(* IEC 61131-3 sources: plc-workbench/outputs/tia_32x4_20261108_results/tasks/15_PUBLIC_03/self_A/details/submissions/1/evaluation/formal, 1 file *)

(* ---- normalized.st ---- *)
FUNCTION_BLOCK Q03

   VAR_INPUT
      Value : REAL;
      hiLevel : REAL;
      loLevel : REAL;
      hystWindow : REAL;
   END_VAR
   VAR_OUTPUT
      hiAlarm : BOOL;
      loAlarm : BOOL;
      error : BOOL;
      status : WORD;
   END_VAR
   VAR
      valid : BOOL;
   END_VAR
VAR_INPUT
WBTEMP_0 : BOOL;
END_VAR

valid := WBTEMP_0;
   // Validity of configuration
   valid := FALSE;

   IF loLevel >= hiLevel THEN
      // Invalid limits: loLevel must be smaller than hiLevel
      error := TRUE;
      status := 16#8001;
   ELSIF hystWindow >= (hiLevel - loLevel) THEN
      // Invalid hysteresis window relative to the deviation range
      error := TRUE;
      status := 16#8002;
   ELSE
      valid := TRUE;
      error := FALSE;
      status := 16#0000;
   END_IF;

   IF valid THEN
      // High alarm with hysteresis
      IF Value > hiLevel THEN
         hiAlarm := TRUE;
      ELSIF Value < (hiLevel - hystWindow) THEN
         hiAlarm := FALSE;
      END_IF;

      // Low alarm with hysteresis
      IF Value < loLevel THEN
         loAlarm := TRUE;
      ELSIF Value > (loLevel + hystWindow) THEN
         loAlarm := FALSE;
      END_IF;
   END_IF;

END_FUNCTION_BLOCK
